TYPE ST_CamXYVA :
STRUCT
	fDx: LREAL;
	fDy: LREAL;
	fDv: LREAL;
	fDa: LREAL;
	fDj: LREAL;
	///Segment TYPE
	nMotionFunctionType: UINT;
END_STRUCT
END_TYPE

(* stored: Version 1.1.0.1, ProductVersion 3.1.4024.12
   DUT ST_CamXYVA: Id {33ff0f9a-99d0-4c23-b6e5-3a97473c97c8} *)
